FUNCTION_BLOCK FB_JSReference
VAR_INPUT
	bStartX	:	BOOL;
	bStartY	:	BOOL;
	bStartZ	:	BOOL;
END_VAR
VAR_OUTPUT
	bReferenced: BOOL := FALSE;
END_VAR
VAR_IN_OUT
	motX:	AXIS_REF;
	motY:	AXIS_REF;
	motZ:	AXIS_REF;
END_VAR	
VAR
	JS_MC_X :	JS_MC_REF;
	JS_MC_Y :	JS_MC_REF;
	JS_MC_Z :	JS_MC_REF;
	Done_X	:	BOOL;
	Done_Y	:	BOOL;
	Done_Z	:	BOOL;
END_VAR

JS_MC_X(
	Axis	:=	motX,
	bExecute:=	bStartX,
	bAbort	:=	FALSE,
	bForceNewRef	:=FALSE,
	iTypeGantry	:=0,
	Done	=>	Done_X);
	
JS_MC_Y(
	Axis	:=	motY,
	bExecute:=	bStartY,
	bAbort	:=	FALSE,
	bForceNewRef	:=FALSE,
	iTypeGantry	:=0,
	Done	=>	Done_Y);
	
JS_MC_Z(
	Axis	:=	motZ,
	bExecute:=	bStartZ,
	bAbort	:=	FALSE,
	bForceNewRef	:=FALSE,
	iTypeGantry	:=0,
	Done	=>	Done_Z);

IF bStartX OR bStartY OR bStartZ THEN
	bReferenced	:=	
		((NOT bStartX) OR Done_X) AND
		((NOT bStartY) OR Done_Y) AND
		((NOT bStartZ) OR Done_Z);
ELSE
	bReferenced	:=	FALSE;
END_IF

END_FUNCTION_BLOCK

(* stored: Version 1.1.0.1, ProductVersion 3.1.4024.15
   POU FB_JSReference: Id {e381aa14-296c-43d4-92a2-46799356c340}, SpecialFunc None *)
